{attribute 'qualified_only'}
  VAR_GLOBAL
  END_VAR

(* stored: Version 1.1.0.1, ProductVersion 3.1.4026.13
   GVL GVL_Inputs: Id {61bea2d8-6613-4ba3-addb-3df0034b2c51} *)
